(* IEC 61131-3 sources: codesys-framework/txt/application/WeVe Visu (library)/Controller, 9 files *)

(* ---- GVL_Color.gvl.st ---- *)
VAR_GLOBAL CONSTANT
	cColorUnknown 					: DWORD 	:= 16#FFCCCCCC;
	cColorNoCarrier 				: DWORD 	:= 16#FFFF0000;
	cColorCarrierWithoutTube 		: DWORD 	:= 16#FFFF8000;
	cColorCarrierWithTube 			: DWORD 	:= 16#FFFFFF00;
	cColorCarrierWithPackage 		: DWORD 	:= 16#00FFFFFF;
	cColorNewCarrier 				: DWORD 	:= 16#FF0000FF;
	cColorActivePosition 			: DWORD 	:= 16#8000FF00;
	cColorNotEnabled 				: DWORD 	:= 16#FF4D4D4D;
	cColorNotPresent 				: DWORD 	:= 16#FF000000;
END_VAR

(* ---- FB_GeneralInputsController.pou.st ---- *)
FUNCTION_BLOCK FB_GeneralInputsController
VAR_INPUT
END_VAR
VAR_OUTPUT
END_VAR
VAR
	_fbUserRequest 			: I_UserRequestModule;
	_fbSignalLamp 			: I_SignalLampModule;
	_fbEmergencyStop 		: I_EmergencyStopModule;

	(* General inputs *)
	_xBtnEmergencyStop 		: BOOL;
	_btnStart 				: FB_VisuButtonTrigger;
	_btnStop 				: FB_VisuButtonTrigger;
	_btnReset 				: FB_VisuButtonTrigger;

	_tonDelayedStop 		: TON;
	_rtrigDelayedStop 		: R_TRIG;

	_xBtnSimulation 		: BOOL;

	_xEmergencyBtnState 	: BOOL;

	_scSignalLamp 			: SC_SignalLamp;
	_xSignalLightStartBtn 	: BOOL;
	_xSignalLightResetBtn 	: BOOL;
	_xSignalLightGreen 		: BOOL;
	_xSignalLightOrange 	: BOOL;
	_xSignalLightRed 		: BOOL;

	_iStopCounter 			: UINT;
	_tonCounter 			: TON;
END_VAR

// --- BEGIN IMPLEMENTATION ---

_btnStart();

IF _btnStart.RQ THEN
	_fbUserRequest.Start(sSource := 'Visu');
END_IF

_btnStop();

IF _btnStop.RQ THEN
	_fbUserRequest.Stop(sSource := 'Visu');
	_iStopCounter := _iStopCounter + 1;
END_IF

_tonCounter(IN := _iStopCounter > 0, PT := T#500MS);

IF _tonCounter.Q THEN
	_iStopCounter := 0;
END_IF

IF _iStopCounter >= 2 THEN
	_fbUserRequest.QuickStop();
END_IF

_tonDelayedStop(IN := _btnStop.State, PT := cStopDelayTime);
_rtrigDelayedStop(CLK := _tonDelayedStop.Q);

IF _rtrigDelayedStop.Q THEN
	_fbUserRequest.ResetSequence(sSource := 'Visu');
END_IF

_btnReset();

IF _btnReset.RQ THEN
	_fbUserRequest.ResetSafety(sSource := 'Visu');
END_IF

_xEmergencyBtnState := FALSE;

IF _fbEmergencyStop.State = E_EmergencyStopState.NOK THEN
	_xEmergencyBtnState := TRUE;
END_IF

_scSignalLamp := _fbSignalLamp.SignalLamp;

_xSignalLightStartBtn 	:= _scSignalLamp.xStartBtn;
_xSignalLightResetBtn 	:= _scSignalLamp.xResetBtn;
_xSignalLightGreen 		:= _scSignalLamp.xGreen;
_xSignalLightOrange 	:= _scSignalLamp.xOrange;
_xSignalLightRed 		:= _scSignalLamp.xRed;

(* ---- FB_JobManagerController.pou.st ---- *)
FUNCTION_BLOCK FB_JobManagerController
VAR_INPUT
END_VAR
VAR_OUTPUT
END_VAR
VAR
	_fbJobSrv 				: I_JobService;

	_eJobType 				: E_JobRequests;
	_scJob 					: SC_JobRequest;

	_ascSrvJobs 			: ARRAY [1..cMaxNbrOfJobs] OF SC_JobRequest;
	_ascJobs 				: ARRAY [1..cMaxNbrOfJobs] OF SC_VisuJobInfo;
	_scEmptyJob 			: SC_VisuJobInfo;

	_i 						: UINT;

END_VAR

// --- BEGIN IMPLEMENTATION ---

_ascSrvJobs := _fbJobSrv.GetJobs();

FOR _i := 1 TO cMaxNbrOfJobs DO

	IF _ascSrvJobs[_i].eState <> E_JobStates.None THEN
		_ascJobs[_i].eJobType 		:= _ascSrvJobs[_i].eType;
		_ascJobs[_i].eJobState 		:= _ascSrvJobs[_i].eState;
		_ascJobs[_i].eJobPriority 	:= _ascSrvJobs[_i].ePriority;
		_ascJobs[_i].eFrame 		:= _ascSrvJobs[_i].scPosition.eStorage;
		_ascJobs[_i].eSide 			:= _ascSrvJobs[_i].scPosition.eSide;
	ELSE
		_ascJobs[_i] := _scEmptyJob;
	END_IF

END_FOR

(* ---- FB_ManualController.pou.st ---- *)
FUNCTION_BLOCK FB_ManualController
VAR_OUTPUT
	xManualMode 			: BOOL;
	xEnabled 				: BOOL;
END_VAR
VAR
	_fbManualMode 			: I_Mode;

	_btnRequestHomePos 			: FB_VisuButtonTrigger;
	_btnCalibrateCamGripper		: FB_VisuButtonTrigger;
	_btnCalibrateCamAngled		: FB_VisuButtonTrigger;
	_btnMeasure 				: FB_VisuButtonTrigger;
	_btnFindCoils				: FB_VisuButtonTrigger;
	_btnPickCoil				: FB_VisuButtonTrigger;
	_btnPickDropCoil			: FB_VisuButtonTrigger;
	_btnRequestTopOfMaster		: FB_VisuButtonTrigger;
	_btnRequestDisable			: FB_VisuButtonTrigger;
	_btnDropCoil				: FB_VisuButtonTrigger;
	_btnDropCoilOnFloor			: FB_VisuButtonTrigger;
	_btnPickTopCoil				: FB_VisuButtonTrigger;
	_btnReleaseBuggy			: FB_VisuButtonTrigger;
	_btnClampBuggy				: FB_VisuButtonTrigger;
	_btnFindAndWait				: FB_VisuButtonTrigger;
	_btnPickDropFromPos			: FB_VisuButtonTrigger;
	_btnPickDropCardboard		: FB_VisuButtonTrigger;
	_btnCheckEmptyLayer			: FB_VisuButtonTrigger;
	_btnCheckEmptyLayerLaser	: FB_VisuButtonTrigger;
	_btnDropCardboard			: FB_VisuButtonTrigger;
	_btnMeasureCoilOrCardboard	: FB_VisuButtonTrigger;
	_btnCheckStorageOrientation	: FB_VisuButtonTrigger;

	_scRobotPosition 		: SC_RobotPosition;

	_scRobotPosRealsTemp	: SC_RobotPositionReals;

	_ascCamJobsToTry		: ARRAY [1..5] OF UINT;

END_VAR

// --- BEGIN IMPLEMENTATION ---

xManualMode := _fbManualMode.Mode = E_DefaultModes.Manual AND _fbManualMode.State = E_ModeStates.StandBy;

_btnRequestHomePos();
IF _btnRequestHomePos.RQ THEN
	_fbManualMode.SetRequest(iRequest := E_JobRequests.ManualHomePosition);
END_IF

_btnCalibrateCamGripper();
IF _btnCalibrateCamGripper.RQ THEN
	_fbManualMode.SetRequest(iRequest := E_JobRequests.ManualCalibrateCamGripper);
END_IF

_btnCalibrateCamAngled();
IF _btnCalibrateCamAngled.RQ THEN
	_fbManualMode.SetRequest(iRequest := E_JobRequests.ManualCalibrateCamAngled);
END_IF

_btnMeasure();
IF _btnMeasure.RQ THEN
	_scRobotPosition.scRobotPosition := PersistentVars.scFeedrobot.RobotArm.MeasurePositionLeft;
	_fbManualMode.SetRequest(iRequest := E_JobRequests.ManualMeasure, pData := ADR(_scRobotPosition), pSize := SIZEOF(_scRobotPosition));
END_IF

_btnFindCoils();
IF _btnFindCoils.RQ THEN
	//set job request
	_fbManualMode.SetRequest(iRequest := E_JobRequests.ManualFindCoils, pData := ADR(_scRobotPosition), pSize := SIZEOF(_scRobotPosition));
END_IF

_btnFindAndWait();
IF _btnFindAndWait.RQ THEN
	//set job request
	_fbManualMode.SetRequest(iRequest := E_JobRequests.ManualFindAndWait, pData := ADR(_scRobotPosition), pSize := SIZEOF(_scRobotPosition));
END_IF

_btnPickCoil();
IF _btnPickCoil.RQ THEN
	//get robot orientation
	_scRobotPosRealsTemp := PersistentVars.scFeedRobot.RobotArm.refPosPickCoils;
	_scRobotPosRealsTemp.posX := _scRobotPosition.scRobotPosition.posX;
	_scRobotPosRealsTemp.posY := _scRobotPosition.scRobotPosition.posY;
	_scRobotPosRealsTemp.posZ := _scRobotPosition.scRobotPosition.posZ;
	_scRobotPosRealsTemp.posRX := _scRobotPosition.scRobotPosition.posRX;
	_scRobotPosRealsTemp.posRY := _scRobotPosition.scRobotPosition.posRY;
	_scRobotPosRealsTemp.posRZ := _scRobotPosition.scRobotPosition.posRZ;
	_scRobotPosRealsTemp.ToolID := _scRobotPosition.scRobotPosition.ToolID;
	//trensfrom to correct buggy side
	_scRobotPosition.scRobotPosition := _scRobotposrealstemp;
	//set job request
	_fbManualMode.SetRequest(iRequest := E_JobRequests.ManualPickCoil, pData := ADR(_scRobotPosition), pSize := SIZEOF(_scRobotPosition));
END_IF

_btnRequestTopOfMaster();
IF _btnRequestTopOfMaster.RQ THEN
	_fbManualMode.SetRequest(iRequest := E_JobRequests.ManualTopOfMaster);
END_IF

_btnRequestDisable();
IF _btnRequestDisable.RQ THEN
	_fbManualMode.SetRequest(iRequest := E_JobRequests.ManualDisable);
END_IF

_btnDropCoil();
IF _btnDropCoil.RQ THEN
	_fbManualMode.SetRequest(iRequest := E_JobRequests.ManualDropCoil,pData := ADR(_scRobotPosition), pSize := SIZEOF(_scRobotPosition));
END_IF

_btnDropCoilOnFloor();
IF _btnDropCoilOnFloor.RQ THEN
	_fbManualMode.SetRequest(iRequest := E_JobRequests.ManualDropFloor);
END_IF

_btnPickTopCoil();
IF _btnPickTopCoil.RQ THEN
	//set job request
	_fbManualMode.SetRequest(iRequest := E_JobRequests.ManualPickTopCoil, pData := ADR(_scRobotPosition), pSize := SIZEOF(_scRobotPosition));
END_IF

_btnReleaseBuggy();
IF _btnReleaseBuggy.RQ THEN
	//set job request
	_fbManualMode.SetRequest(iRequest := E_JobRequests.ManualReleaseBuggy, pData := ADR(_scRobotPosition), pSize := SIZEOF(_scRobotPosition));
END_IF

_btnClampBuggy();
IF _btnClampBuggy.RQ THEN
	//set job request
	_fbManualMode.SetRequest(iRequest := E_JobRequests.ManualClampBuggy, pData := ADR(_scRobotPosition), pSize := SIZEOF(_scRobotPosition));
END_IF

_btnPickDropCoil();
IF _btnPickDropCoil.RQ THEN
	//set job request
	_fbManualMode.SetRequest(iRequest := E_JobRequests.ManualPickDropCoil, pData := ADR(_scRobotPosition), pSize := SIZEOF(_scRobotPosition));
END_IF

_btnPickDropFromPos();
IF _btnPickDropFromPos.RQ THEN
	//set job request
	_fbManualMode.SetRequest(iRequest := E_JobRequests.ManualPickDropFromPos, pData := ADR(_scRobotPosition), pSize := SIZEOF(_scRobotPosition));
END_IF

_btnPickDropCardboard();
IF _btnPickDropCardboard.RQ THEN
	//set job request
	_fbManualMode.SetRequest(iRequest := E_JobRequests.ManualPickDropCardboard, pData := ADR(_scRobotPosition), pSize := SIZEOF(_scRobotPosition));
END_IF

_btnCheckEmptyLayer();
IF _btnCheckEmptyLayer.RQ THEN
	//set job request
	_fbManualMode.SetRequest(iRequest := E_JobRequests.ManualCheckEmptyLayer, pData := ADR(_scRobotPosition), pSize := SIZEOF(_scRobotPosition));
END_IF

_btnCheckEmptyLayerLaser();
IF _btnCheckEmptyLayerLaser.RQ THEN
	//set job request
	_fbManualMode.SetRequest(iRequest := E_JobRequests.ManualCheckEmptyLayerLaser, pData := ADR(_scRobotPosition), pSize := SIZEOF(_scRobotPosition));
END_IF

_btnDropCardboard();
IF _btnDropCardboard.RQ THEN
	_fbManualMode.SetRequest(iRequest := E_JobRequests.ManualDropCardboard, pData := ADR(_scRobotPosition), pSize := SIZEOF(_scRobotPosition));
END_IF

_btnMeasureCoilOrCardboard();
IF _btnMeasureCoilOrCardboard.RQ THEN
	_scRobotPosition.scRobotPosition := PersistentVars.scFeedrobot.RobotArm.MeasurePositionLeft;
	_fbManualMode.SetRequest(iRequest := E_JobRequests.ManualMeasureCoilOrCardboard, pData := ADR(_scRobotPosition), pSize := SIZEOF(_scRobotPosition));
END_IF

_btnCheckStorageOrientation();
IF _btnCheckStorageOrientation.RQ THEN
	_scRobotPosition.scRobotPosition := PersistentVars.scFeedrobot.RobotArm.MeasurePositionCheckOrientation;
	_fbManualMode.SetRequest(iRequest := E_JobRequests.ManualCheckStorageOrientation, pData := ADR(_scRobotPosition), pSize := SIZEOF(_scRobotPosition));
END_IF

(* ---- FB_ModeController.pou.st ---- *)
FUNCTION_BLOCK FB_ModeController
VAR_INPUT
	pOpModeSrv 				: POINTER TO FB_ModeService;
END_VAR
VAR_OUTPUT
END_VAR
VAR
	_fbOpModeSrv 			: I_ModeService;
	_fbLogger 				: I_EventHandlerService;

	_btnRequestAutomatic 	: FB_VisuButtonTrigger;
	_btnRequestManual 		: FB_VisuButtonTrigger;
	_btnRequestMaintenance 	: FB_VisuButtonTrigger;
	_btnRequestTest 		: FB_VisuButtonTrigger;

	_ascMessages 			: ARRAY[1..cNbrOfLogMessages] OF SC_LogMessage;
END_VAR

// --- BEGIN IMPLEMENTATION ---

_btnRequestAutomatic();
_btnRequestManual();
_btnRequestMaintenance();
_btnRequestTest();

IF _btnRequestAutomatic.RQ THEN
	_fbOpModeSrv.RequestMode(eMode := E_DefaultModes.Auto);
END_IF

IF _btnRequestManual.RQ THEN
	_fbOpModeSrv.RequestMode(eMode := E_DefaultModes.Manual);
END_IF

IF _btnRequestMaintenance.RQ THEN
	_fbOpModeSrv.RequestMode(eMode := E_DefaultModes.Maintenance);
END_IF

IF _btnRequestTest.RQ THEN
	_fbOpModeSrv.RequestMode(eMode := E_DefaultModes.UserDefined1);
END_IF

_ascMessages := _fbLogger.GetMessages();

(* ---- FB_NavBarController.pou.st ---- *)
FUNCTION_BLOCK FB_NavBarController
VAR_INPUT
	xHoverParameters 			: BOOL;
END_VAR
VAR_OUTPUT
	iFrame 						: UINT;
	xHideParameters 			: BOOL;
END_VAR
VAR
	_btnOperationalMode 		: FB_VisuButtonTrigger;

	_btnParameters 				: FB_VisuButtonTrigger;
	_btnSysParFR 				: FB_VisuButtonTrigger;
	_btnSysParBuggy 			: FB_VisuButtonTrigger;
	_btnSysParSafety 			: FB_VisuButtonTrigger;

	_btnJobManager 				: FB_VisuButtonTrigger;
	_btnManualRequest 			: FB_VisuButtonTrigger;
	_btnFeedRobot 				: FB_VisuButtonTrigger;
	_btnYarnStorage 			: FB_VisuButtonTrigger;

	_tonHideParameters 			: TON;
	_rtrigHideParameters 		: R_TRIG;
END_VAR

// --- BEGIN IMPLEMENTATION ---

ProcessFBs();
HandleButtonClicks();

IF _btnParameters.RQ THEN
	xHideParameters := NOT xHideParameters;
END_IF

_tonHideParameters(IN := NOT xHoverParameters, PT := T#250MS);
_rtrigHideParameters(CLK := _tonHideParameters.Q);

IF _rtrigHideParameters.Q THEN
	xHideParameters := TRUE;
END_IF

(* ---- FB_ParametersController.pou.st ---- *)
FUNCTION_BLOCK FB_ParametersController
VAR_INPUT
END_VAR
VAR_OUTPUT
END_VAR
VAR
	_fbParameterSrv 			: I_ParameterService;

	_btnLoadDefaultParameters 	: FB_VisuButtonTrigger;
	_aiNumber 					: ARRAY[1..3] OF INT := [1,2,3];
END_VAR

// --- BEGIN IMPLEMENTATION ---

_btnLoadDefaultParameters();

IF _btnLoadDefaultParameters.RQ THEN
	_fbParameterSrv.LoadDefaultRecipeSettings();
	_fbParameterSrv.LoadDefaultSystemSettings();
END_IF

(* ---- FB_VisuButtonTrigger.pou.st ---- *)
FUNCTION_BLOCK FB_VisuButtonTrigger
VAR_INPUT
	xbtn 		: BOOL;
END_VAR
VAR_OUTPUT
	RQ 			: BOOL;
	FQ 			: BOOL;
	State 		: BOOL;
END_VAR
VAR
	_rtrigger 	: R_TRIG;
	_ftrigger 	: F_TRIG;
END_VAR

// --- BEGIN IMPLEMENTATION ---

State := xbtn;

_rtrigger(CLK := xbtn, Q => RQ);
_ftrigger(CLK := xbtn, Q => FQ);

(* ---- FB_YarnStorageController.pou.st ---- *)
FUNCTION_BLOCK FB_YarnStorageController
VAR_INPUT
END_VAR
VAR_OUTPUT
END_VAR
VAR
	_fbYarnStorageSrv 			: I_YarnStorageService;

	_btnClearStorage 			: FB_VisuButtonTrigger;
	_btnNewPallet				: FB_VisuButtonTrigger;
	_fbStorage 					: I_YarnStorageModule;

	_iStorage 					: E_UserFrame;
	_aState 					: ARRAY[1..2] OF E_StorageState;
	_NbrOfCoilsBase				: UINT;
	_NbrOfCoilsInverted			: UINT;
	_ascCoilPositionsBase		: ARRAY [0..cMaxNbrCoilPositions] OF SC_RobotPositionReals;
	_ascCoilPositionsInverted	: ARRAY [0..cMaxNbrCoilPositions] OF SC_RobotPositionReals;

END_VAR

// --- BEGIN IMPLEMENTATION ---

IF _iStorage < 1 OR _iStorage > 8 THEN
	_iStorage := 1;
END_IF

_aState := _fbYarnStorageSrv.GetStates(_iStorage);

_NbrOfCoilsBase		:= _fbYarnStorageSrv.NbrOfCoils(eStorage := _iStorage, eSide := E_FrameSide.Base);
//_NbrOfCoilsInverted :=_fbYarnStorageSrv.NbrOfCoils(eStorage := _iStorage, eSide := E_FrameSide.Inverted);

_ascCoilPositionsBase := _fbYarnStorageSrv.GetRobotPositions(eStorage := _iStorage, eSide := E_FrameSide.Base);
//_ascCoilPositionsInverted := _fbYarnStorageSrv.GetRobotPositions(eStorage := _iStorage, eSide := E_FrameSide.Inverted);

_btnClearStorage();
IF _btnClearStorage.RQ THEN
	_fbStorage := _fbYarnStorageSrv.GetStorage(id := _iStorage);
	_fbStorage.SetSideState(eSide := 1, eState := E_StorageState.New);
	_fbStorage.SetSideState(eSide := 2, eState := E_StorageState.New);
	_fbStorage.ResetData();
END_IF

_btnNewPallet();
IF _btnNewPallet.RQ THEN
	_fbStorage := _fbYarnStorageSrv.GetStorage(id := _iStorage);
	_fbStorage.SetSideState(eSide := 1, eState := E_StorageState.New);
	_fbStorage.SetSideState(eSide := 2, eState := E_StorageState.New);
	_fbStorage.ResetData();
END_IF
